FUNCTION_BLOCK MinutesSinceLastAerateBasic (* Basic Function Block Type *)
  (* Standard: 61499-2 *)
  (* Version 0.0, 7/5/2026, Schneider Electric, Template *)
  PACKAGE SE.Nereda;
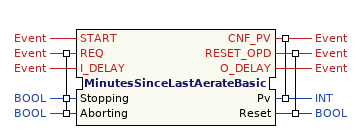
  EVENT_INPUT
    START;
    REQ WITH Stopping, Aborting; (* Normal Execution Request *)
    I_DELAY;
  END_EVENT
  EVENT_OUTPUT
    CNF_PV WITH Pv; (* Execution Confirmation *)
    RESET_OPD WITH Reset;
    O_DELAY;
  END_EVENT
  VAR_INPUT
    Stopping : BOOL;
    Aborting : BOOL;
  END_VAR
  VAR_OUTPUT
    Pv : INT; (* Output event qualifier *)
    Reset : BOOL;
  END_VAR
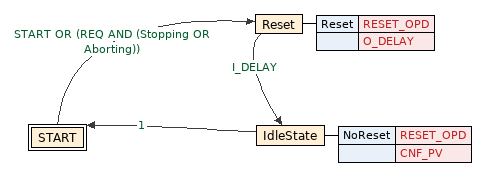
  EC_STATES
    START; (* Initial State *)
    Reset : Reset -> RESET_OPD, -> O_DELAY;
    IdleState : NoReset -> RESET_OPD, -> CNF_PV;
  END_STATES
  EC_TRANSITIONS
    START TO Reset := START OR (REQ AND (Stopping OR Aborting));
    Reset TO IdleState := I_DELAY;
    IdleState TO START := 1;
  END_TRANSITIONS
  ALGORITHM Reset IN ST:
;
Reset := TRUE;
  END_ALGORITHM
  ALGORITHM NoReset IN ST:
;
Pv := 1;
Reset := FALSE;
  END_ALGORITHM
END_FUNCTION_BLOCK
